// --- Siemens Structured Format ---
DATA_BLOCK "model__HS8_IW50_"
{ S7_Optimized_Access := 'TRUE' }
VERSION :
NON_RETAIN
   VAR
      W_i : ARRAY[0..7, 0..39] OF REAL;
      W_f : ARRAY[0..7, 0..39] OF REAL;
      W_g : ARRAY[0..7, 0..39] OF REAL;
      W_o : ARRAY[0..7, 0..39] OF REAL;
      R_i : ARRAY[0..7, 0..7] OF REAL;
      R_f : ARRAY[0..7, 0..7] OF REAL;
      R_g : ARRAY[0..7, 0..7] OF REAL;
      R_o : ARRAY[0..7, 0..7] OF REAL;
      B_i : ARRAY[0..7] OF REAL;
      B_f : ARRAY[0..7] OF REAL;
      B_g : ARRAY[0..7] OF REAL;
      B_o : ARRAY[0..7] OF REAL;
      FC_W : ARRAY[0..39, 0..7] OF REAL;
      FC_B : ARRAY[0..39] OF REAL;
   END_VAR
BEGIN

      W_i[0,0] := 0.02461717;
      W_i[0,1] := 0.08401545;
      W_i[0,2] := -0.12303820;
      W_i[0,3] := -0.02682650;
      W_i[0,4] := 0.14538512;
      W_i[0,5] := 0.05910228;
      W_i[0,6] := -0.06121323;
      W_i[0,7] := 0.19529903;
      W_i[0,8] := 0.21199454;
      W_i[0,9] := -0.29979098;
      W_i[0,10] := -0.09429822;
      W_i[0,11] := -0.28532824;
      W_i[0,12] := 0.06377743;
      W_i[0,13] := -0.06364888;
      W_i[0,14] := 0.00534459;
      W_i[0,15] := 0.03598412;
      W_i[0,16] := 0.04236616;
      W_i[0,17] := 0.00850482;
      W_i[0,18] := 0.00358703;
      W_i[0,19] := 0.18395557;
      W_i[0,20] := 0.05710260;
      W_i[0,21] := 0.31176916;
      W_i[0,22] := 0.17010060;
      W_i[0,23] := -0.01221133;
      W_i[0,24] := -0.19286193;
      W_i[0,25] := -0.07674938;
      W_i[0,26] := -0.40142074;
      W_i[0,27] := -0.50435519;
      W_i[0,28] := 0.04934237;
      W_i[0,29] := -0.24499206;
      W_i[0,30] := 0.63579166;
      W_i[0,31] := -0.13499857;
      W_i[0,32] := 0.02890123;
      W_i[0,33] := -0.00438442;
      W_i[0,34] := -0.02304220;
      W_i[0,35] := -0.28221473;
      W_i[0,36] := -0.00601982;
      W_i[0,37] := -0.39292136;
      W_i[0,38] := -0.02013459;
      W_i[0,39] := -0.00859181;
      W_i[1,0] := -0.17783616;
      W_i[1,1] := 0.10906062;
      W_i[1,2] := 0.27302170;
      W_i[1,3] := 0.03857158;
      W_i[1,4] := 0.15132146;
      W_i[1,5] := -0.07943013;
      W_i[1,6] := -0.12445311;
      W_i[1,7] := 0.10142804;
      W_i[1,8] := 0.17782561;
      W_i[1,9] := -0.34472182;
      W_i[1,10] := -0.15930130;
      W_i[1,11] := 0.11785957;
      W_i[1,12] := 0.12351760;
      W_i[1,13] := 0.01896391;
      W_i[1,14] := -0.06655354;
      W_i[1,15] := 0.10417320;
      W_i[1,16] := 0.02300226;
      W_i[1,17] := -0.06141837;
      W_i[1,18] := 0.28663757;
      W_i[1,19] := -0.05906216;
      W_i[1,20] := -0.01470305;
      W_i[1,21] := 0.12249159;
      W_i[1,22] := 0.08935670;
      W_i[1,23] := -0.19675028;
      W_i[1,24] := 0.48150146;
      W_i[1,25] := 0.29962191;
      W_i[1,26] := 0.04253698;
      W_i[1,27] := -0.01234774;
      W_i[1,28] := -0.20131898;
      W_i[1,29] := -0.28958127;
      W_i[1,30] := 0.30615368;
      W_i[1,31] := -0.00297963;
      W_i[1,32] := 0.24898766;
      W_i[1,33] := -0.17079352;
      W_i[1,34] := -0.01789305;
      W_i[1,35] := -0.07885017;
      W_i[1,36] := 0.02689386;
      W_i[1,37] := 0.36441922;
      W_i[1,38] := -0.06345996;
      W_i[1,39] := 0.09888364;
      W_i[2,0] := 0.10794700;
      W_i[2,1] := 0.01449859;
      W_i[2,2] := 0.11232290;
      W_i[2,3] := 0.04600843;
      W_i[2,4] := 0.15555517;
      W_i[2,5] := -0.08419870;
      W_i[2,6] := 0.10784180;
      W_i[2,7] := -0.13110802;
      W_i[2,8] := 0.01003856;
      W_i[2,9] := 0.13528554;
      W_i[2,10] := -0.08593279;
      W_i[2,11] := 0.15705661;
      W_i[2,12] := 0.00744481;
      W_i[2,13] := 0.14232995;
      W_i[2,14] := -0.07310586;
      W_i[2,15] := 0.11869515;
      W_i[2,16] := 0.16272350;
      W_i[2,17] := 0.01258006;
      W_i[2,18] := 0.17897964;
      W_i[2,19] := -0.08531563;
      W_i[2,20] := -0.06869420;
      W_i[2,21] := -0.05605607;
      W_i[2,22] := -0.24934621;
      W_i[2,23] := 0.02436493;
      W_i[2,24] := 0.04889333;
      W_i[2,25] := -0.20094825;
      W_i[2,26] := -0.40725628;
      W_i[2,27] := -0.16053441;
      W_i[2,28] := -0.17641398;
      W_i[2,29] := -0.18513416;
      W_i[2,30] := 0.09812243;
      W_i[2,31] := -0.24586804;
      W_i[2,32] := 0.18386346;
      W_i[2,33] := -0.37200448;
      W_i[2,34] := -0.30738470;
      W_i[2,35] := 0.07613509;
      W_i[2,36] := -0.04531293;
      W_i[2,37] := -0.08632755;
      W_i[2,38] := -0.13347539;
      W_i[2,39] := -0.03515237;
      W_i[3,0] := -0.04817922;
      W_i[3,1] := -0.16765678;
      W_i[3,2] := -0.00308369;
      W_i[3,3] := -0.41362956;
      W_i[3,4] := -0.07394656;
      W_i[3,5] := 0.09627691;
      W_i[3,6] := 0.11941688;
      W_i[3,7] := -0.17643057;
      W_i[3,8] := 0.06146013;
      W_i[3,9] := 0.13595612;
      W_i[3,10] := 0.21689560;
      W_i[3,11] := 0.08097983;
      W_i[3,12] := -0.05968216;
      W_i[3,13] := 0.06028462;
      W_i[3,14] := -0.33660558;
      W_i[3,15] := -0.14613369;
      W_i[3,16] := 0.15110187;
      W_i[3,17] := 0.02597690;
      W_i[3,18] := 0.00098816;
      W_i[3,19] := 0.26554033;
      W_i[3,20] := 0.06123941;
      W_i[3,21] := -0.20589893;
      W_i[3,22] := -0.01046670;
      W_i[3,23] := -0.35783783;
      W_i[3,24] := -0.18957515;
      W_i[3,25] := -0.03140980;
      W_i[3,26] := 0.00826861;
      W_i[3,27] := 0.05130741;
      W_i[3,28] := 0.13812958;
      W_i[3,29] := -0.19599199;
      W_i[3,30] := -0.16747603;
      W_i[3,31] := -0.13670678;
      W_i[3,32] := -0.15334715;
      W_i[3,33] := -0.32899481;
      W_i[3,34] := 0.07909799;
      W_i[3,35] := -0.27765223;
      W_i[3,36] := -0.03015585;
      W_i[3,37] := 0.07159591;
      W_i[3,38] := -0.33855185;
      W_i[3,39] := -0.69761050;
      W_i[4,0] := 0.10504181;
      W_i[4,1] := 0.00682971;
      W_i[4,2] := -0.05512364;
      W_i[4,3] := -0.42238507;
      W_i[4,4] := 0.21000206;
      W_i[4,5] := 0.08828816;
      W_i[4,6] := -0.25787413;
      W_i[4,7] := 0.18548162;
      W_i[4,8] := 0.07325415;
      W_i[4,9] := -0.16746196;
      W_i[4,10] := -0.23054802;
      W_i[4,11] := -0.17278661;
      W_i[4,12] := 0.19685929;
      W_i[4,13] := -0.06621253;
      W_i[4,14] := -0.04979985;
      W_i[4,15] := -0.02534566;
      W_i[4,16] := -0.05196558;
      W_i[4,17] := -0.02844546;
      W_i[4,18] := 0.21438381;
      W_i[4,19] := -0.22215076;
      W_i[4,20] := 0.01178194;
      W_i[4,21] := -0.06624336;
      W_i[4,22] := -0.05115673;
      W_i[4,23] := -0.23732296;
      W_i[4,24] := -0.09036870;
      W_i[4,25] := -0.09140033;
      W_i[4,26] := 0.12307051;
      W_i[4,27] := -0.02017660;
      W_i[4,28] := -0.07642211;
      W_i[4,29] := -0.01614011;
      W_i[4,30] := -0.17466348;
      W_i[4,31] := -0.15838575;
      W_i[4,32] := 0.18079966;
      W_i[4,33] := 0.33373138;
      W_i[4,34] := 0.09327173;
      W_i[4,35] := -0.13638979;
      W_i[4,36] := -0.08043678;
      W_i[4,37] := -0.09420969;
      W_i[4,38] := -0.03976285;
      W_i[4,39] := 0.22526605;
      W_i[5,0] := 0.46471885;
      W_i[5,1] := 0.24254853;
      W_i[5,2] := -0.00896330;
      W_i[5,3] := -0.40931293;
      W_i[5,4] := 0.07764716;
      W_i[5,5] := -0.12571707;
      W_i[5,6] := -0.07207277;
      W_i[5,7] := -0.58136684;
      W_i[5,8] := -0.70827621;
      W_i[5,9] := 0.13912673;
      W_i[5,10] := 0.00305168;
      W_i[5,11] := 0.10330518;
      W_i[5,12] := -0.39406857;
      W_i[5,13] := -0.13641670;
      W_i[5,14] := -0.13437758;
      W_i[5,15] := 0.32282859;
      W_i[5,16] := 0.14888868;
      W_i[5,17] := 0.07580157;
      W_i[5,18] := 0.78602076;
      W_i[5,19] := -0.46361649;
      W_i[5,20] := -0.12363275;
      W_i[5,21] := 0.16991106;
      W_i[5,22] := -0.08441558;
      W_i[5,23] := 0.01862625;
      W_i[5,24] := 0.45371729;
      W_i[5,25] := 1.03232503;
      W_i[5,26] := 0.00888214;
      W_i[5,27] := -0.04149527;
      W_i[5,28] := -0.06423787;
      W_i[5,29] := -0.13104723;
      W_i[5,30] := -0.16760458;
      W_i[5,31] := -0.06425823;
      W_i[5,32] := 0.11957818;
      W_i[5,33] := 0.10409375;
      W_i[5,34] := 0.68515724;
      W_i[5,35] := 0.21046008;
      W_i[5,36] := 0.09369295;
      W_i[5,37] := -0.08919100;
      W_i[5,38] := -0.09835245;
      W_i[5,39] := 0.00684949;
      W_i[6,0] := 0.04514975;
      W_i[6,1] := -0.18210933;
      W_i[6,2] := -0.00654514;
      W_i[6,3] := -0.41125798;
      W_i[6,4] := 0.04396775;
      W_i[6,5] := -0.00702968;
      W_i[6,6] := -0.05002901;
      W_i[6,7] := -0.03861308;
      W_i[6,8] := 0.06189432;
      W_i[6,9] := -0.02187389;
      W_i[6,10] := 0.03767673;
      W_i[6,11] := -0.55604023;
      W_i[6,12] := -0.48857787;
      W_i[6,13] := 0.13115734;
      W_i[6,14] := -0.05613643;
      W_i[6,15] := -0.11288932;
      W_i[6,16] := 0.17460676;
      W_i[6,17] := -0.26465502;
      W_i[6,18] := 0.16549894;
      W_i[6,19] := 0.29697806;
      W_i[6,20] := 0.23571719;
      W_i[6,21] := -0.09589785;
      W_i[6,22] := 0.59926170;
      W_i[6,23] := -0.08488554;
      W_i[6,24] := 0.70308256;
      W_i[6,25] := 0.90409851;
      W_i[6,26] := -0.01121288;
      W_i[6,27] := -0.09806376;
      W_i[6,28] := -0.02374482;
      W_i[6,29] := -0.20431902;
      W_i[6,30] := 0.48442781;
      W_i[6,31] := -0.11867638;
      W_i[6,32] := 0.28192973;
      W_i[6,33] := 0.13702093;
      W_i[6,34] := 0.91159022;
      W_i[6,35] := -0.05850424;
      W_i[6,36] := -0.02443852;
      W_i[6,37] := 0.08158594;
      W_i[6,38] := -0.16384257;
      W_i[6,39] := 0.04486246;
      W_i[7,0] := -0.16619515;
      W_i[7,1] := -0.08064937;
      W_i[7,2] := 0.17380525;
      W_i[7,3] := -0.35741210;
      W_i[7,4] := 0.25576842;
      W_i[7,5] := -0.11047508;
      W_i[7,6] := -0.00358257;
      W_i[7,7] := 0.22714809;
      W_i[7,8] := 0.14583488;
      W_i[7,9] := -0.14972806;
      W_i[7,10] := -0.14519584;
      W_i[7,11] := -0.41559315;
      W_i[7,12] := -0.01696615;
      W_i[7,13] := -0.28414848;
      W_i[7,14] := 0.06566004;
      W_i[7,15] := 0.09450804;
      W_i[7,16] := -0.03949518;
      W_i[7,17] := 0.04709280;
      W_i[7,18] := 0.19348225;
      W_i[7,19] := 0.10500827;
      W_i[7,20] := -0.09005301;
      W_i[7,21] := -0.34911180;
      W_i[7,22] := -0.00604367;
      W_i[7,23] := -0.15790336;
      W_i[7,24] := 0.51519841;
      W_i[7,25] := 1.09936786;
      W_i[7,26] := -0.23214035;
      W_i[7,27] := -0.30644259;
      W_i[7,28] := 0.08868466;
      W_i[7,29] := 0.18681195;
      W_i[7,30] := 0.44118169;
      W_i[7,31] := 0.16998404;
      W_i[7,32] := -0.39800110;
      W_i[7,33] := 0.02014814;
      W_i[7,34] := 0.50454497;
      W_i[7,35] := -0.04675045;
      W_i[7,36] := -0.05744690;
      W_i[7,37] := 0.17443271;
      W_i[7,38] := -0.05675455;
      W_i[7,39] := 0.18483149;
      W_f[0,0] := -0.08831103;
      W_f[0,1] := 0.00681163;
      W_f[0,2] := -0.02927266;
      W_f[0,3] := 0.05481192;
      W_f[0,4] := -0.06411999;
      W_f[0,5] := 0.00323826;
      W_f[0,6] := 0.04202358;
      W_f[0,7] := -0.14036146;
      W_f[0,8] := -0.12626842;
      W_f[0,9] := 0.10009770;
      W_f[0,10] := 0.02791548;
      W_f[0,11] := -0.04096280;
      W_f[0,12] := -0.00354303;
      W_f[0,13] := 0.01158499;
      W_f[0,14] := -0.04464640;
      W_f[0,15] := -0.08357976;
      W_f[0,16] := 0.04911109;
      W_f[0,17] := 0.09140756;
      W_f[0,18] := -0.03252059;
      W_f[0,19] := 0.01830712;
      W_f[0,20] := 0.01689613;
      W_f[0,21] := 0.22018659;
      W_f[0,22] := 0.08402620;
      W_f[0,23] := -0.07398796;
      W_f[0,24] := 0.08441300;
      W_f[0,25] := 0.18096766;
      W_f[0,26] := 0.05508868;
      W_f[0,27] := -0.13029598;
      W_f[0,28] := -0.02453627;
      W_f[0,29] := 0.12306897;
      W_f[0,30] := 0.37074596;
      W_f[0,31] := 0.04067184;
      W_f[0,32] := 0.33210105;
      W_f[0,33] := 0.17263570;
      W_f[0,34] := 0.02185974;
      W_f[0,35] := 0.21439323;
      W_f[0,36] := 0.00803035;
      W_f[0,37] := 0.09185252;
      W_f[0,38] := -0.03025025;
      W_f[0,39] := 0.16901997;
      W_f[1,0] := -0.08017771;
      W_f[1,1] := 0.05072340;
      W_f[1,2] := -0.15171054;
      W_f[1,3] := -0.04507771;
      W_f[1,4] := -0.01952654;
      W_f[1,5] := 0.01524715;
      W_f[1,6] := -0.03147047;
      W_f[1,7] := -0.02802088;
      W_f[1,8] := -0.15045448;
      W_f[1,9] := 0.13191310;
      W_f[1,10] := 0.00395375;
      W_f[1,11] := -0.03943809;
      W_f[1,12] := -0.13766901;
      W_f[1,13] := -0.04960233;
      W_f[1,14] := -0.11882943;
      W_f[1,15] := -0.18921053;
      W_f[1,16] := 0.07628337;
      W_f[1,17] := -0.01504870;
      W_f[1,18] := 0.23253591;
      W_f[1,19] := 0.00738192;
      W_f[1,20] := 0.02966039;
      W_f[1,21] := -0.07575663;
      W_f[1,22] := 0.28070211;
      W_f[1,23] := 0.04504234;
      W_f[1,24] := 0.44733906;
      W_f[1,25] := 0.76406956;
      W_f[1,26] := -0.18153259;
      W_f[1,27] := -0.01630468;
      W_f[1,28] := 0.04244527;
      W_f[1,29] := -0.03562038;
      W_f[1,30] := 0.06799272;
      W_f[1,31] := -0.07704592;
      W_f[1,32] := 0.08059093;
      W_f[1,33] := 0.21711972;
      W_f[1,34] := 0.58922273;
      W_f[1,35] := -0.24995837;
      W_f[1,36] := -0.01296289;
      W_f[1,37] := -0.02005322;
      W_f[1,38] := 0.11887441;
      W_f[1,39] := 0.13964133;
      W_f[2,0] := 0.02022752;
      W_f[2,1] := -0.03258032;
      W_f[2,2] := 0.02105030;
      W_f[2,3] := -0.01033732;
      W_f[2,4] := -0.02927784;
      W_f[2,5] := 0.05956579;
      W_f[2,6] := -0.06668916;
      W_f[2,7] := -0.06423724;
      W_f[2,8] := -0.06636658;
      W_f[2,9] := 0.16499053;
      W_f[2,10] := -0.01066389;
      W_f[2,11] := -0.08655350;
      W_f[2,12] := 0.03831896;
      W_f[2,13] := 0.02458346;
      W_f[2,14] := 0.12203392;
      W_f[2,15] := -0.07686506;
      W_f[2,16] := -0.09261417;
      W_f[2,17] := -0.01410419;
      W_f[2,18] := 0.05016823;
      W_f[2,19] := -0.13551356;
      W_f[2,20] := 0.00147612;
      W_f[2,21] := -0.01080879;
      W_f[2,22] := -0.23093474;
      W_f[2,23] := 0.18362746;
      W_f[2,24] := 0.34206459;
      W_f[2,25] := 0.11531623;
      W_f[2,26] := -0.10813569;
      W_f[2,27] := -0.03727976;
      W_f[2,28] := 0.08597951;
      W_f[2,29] := 0.16925062;
      W_f[2,30] := 0.14001821;
      W_f[2,31] := 0.08336479;
      W_f[2,32] := -0.13725568;
      W_f[2,33] := 0.14078599;
      W_f[2,34] := -0.22189134;
      W_f[2,35] := 0.07339284;
      W_f[2,36] := 0.01494332;
      W_f[2,37] := -0.16808337;
      W_f[2,38] := 0.02411579;
      W_f[2,39] := 0.21152344;
      W_f[3,0] := -0.03794771;
      W_f[3,1] := 0.05475021;
      W_f[3,2] := -0.02614000;
      W_f[3,3] := 0.08930103;
      W_f[3,4] := 0.04492093;
      W_f[3,5] := 0.03020424;
      W_f[3,6] := -0.07041149;
      W_f[3,7] := 0.23536491;
      W_f[3,8] := -0.04178810;
      W_f[3,9] := -0.19159153;
      W_f[3,10] := -0.06868339;
      W_f[3,11] := -0.16539882;
      W_f[3,12] := 0.12754864;
      W_f[3,13] := -0.13497283;
      W_f[3,14] := 0.13930795;
      W_f[3,15] := 0.00134255;
      W_f[3,16] := -0.03635018;
      W_f[3,17] := 0.02573154;
      W_f[3,18] := -0.41695386;
      W_f[3,19] := -0.18809830;
      W_f[3,20] := 0.04352702;
      W_f[3,21] := 0.16437882;
      W_f[3,22] := 0.06266205;
      W_f[3,23] := 0.08159398;
      W_f[3,24] := 0.04201810;
      W_f[3,25] := -0.19031751;
      W_f[3,26] := -0.17173289;
      W_f[3,27] := -0.23532763;
      W_f[3,28] := 0.17517763;
      W_f[3,29] := 0.39156693;
      W_f[3,30] := 0.25430456;
      W_f[3,31] := 0.07574216;
      W_f[3,32] := 0.27996075;
      W_f[3,33] := 0.00114326;
      W_f[3,34] := -0.28795609;
      W_f[3,35] := 0.19662365;
      W_f[3,36] := 0.02395431;
      W_f[3,37] := -0.22338727;
      W_f[3,38] := 0.15306281;
      W_f[3,39] := 0.18428560;
      W_f[4,0] := 0.01311270;
      W_f[4,1] := -0.01359527;
      W_f[4,2] := -0.03426387;
      W_f[4,3] := -0.05035185;
      W_f[4,4] := 0.09912422;
      W_f[4,5] := -0.04895325;
      W_f[4,6] := -0.03395505;
      W_f[4,7] := -0.02843624;
      W_f[4,8] := -0.08145776;
      W_f[4,9] := 0.08917268;
      W_f[4,10] := -0.00391436;
      W_f[4,11] := -0.07863925;
      W_f[4,12] := 0.03092329;
      W_f[4,13] := 0.01714266;
      W_f[4,14] := -0.03228388;
      W_f[4,15] := -0.05111328;
      W_f[4,16] := 0.02532922;
      W_f[4,17] := -0.04550080;
      W_f[4,18] := -0.03456742;
      W_f[4,19] := -0.02089478;
      W_f[4,20] := 0.09678645;
      W_f[4,21] := -0.08640780;
      W_f[4,22] := 0.02293069;
      W_f[4,23] := 0.05295998;
      W_f[4,24] := 0.11747785;
      W_f[4,25] := 0.00186043;
      W_f[4,26] := -0.20221773;
      W_f[4,27] := -0.01488341;
      W_f[4,28] := 0.04745471;
      W_f[4,29] := -0.16965286;
      W_f[4,30] := 0.02288965;
      W_f[4,31] := -0.03804171;
      W_f[4,32] := 0.13254493;
      W_f[4,33] := -0.13787529;
      W_f[4,34] := -0.43391764;
      W_f[4,35] := -0.24835001;
      W_f[4,36] := 0.07141465;
      W_f[4,37] := -0.29939890;
      W_f[4,38] := -0.01851079;
      W_f[4,39] := 0.08986987;
      W_f[5,0] := -0.14319988;
      W_f[5,1] := -0.10292582;
      W_f[5,2] := -0.17382213;
      W_f[5,3] := -0.01608473;
      W_f[5,4] := -0.00378885;
      W_f[5,5] := 0.00846169;
      W_f[5,6] := 0.06387471;
      W_f[5,7] := 0.20796628;
      W_f[5,8] := -0.42914653;
      W_f[5,9] := 0.01919760;
      W_f[5,10] := 0.04385304;
      W_f[5,11] := 0.01982332;
      W_f[5,12] := 0.11683133;
      W_f[5,13] := 0.07871818;
      W_f[5,14] := -0.12016966;
      W_f[5,15] := -0.06522254;
      W_f[5,16] := -0.10883621;
      W_f[5,17] := -0.02835156;
      W_f[5,18] := -0.26717833;
      W_f[5,19] := 0.08458684;
      W_f[5,20] := -0.00364884;
      W_f[5,21] := -0.04485849;
      W_f[5,22] := -0.19082835;
      W_f[5,23] := 0.06622007;
      W_f[5,24] := 0.45456037;
      W_f[5,25] := 0.15541779;
      W_f[5,26] := 0.00758505;
      W_f[5,27] := 0.07440008;
      W_f[5,28] := 0.05810034;
      W_f[5,29] := 0.14797372;
      W_f[5,30] := -0.11548296;
      W_f[5,31] := 0.02787589;
      W_f[5,32] := -0.27752876;
      W_f[5,33] := -0.08107541;
      W_f[5,34] := -0.09626248;
      W_f[5,35] := -0.23543228;
      W_f[5,36] := -0.00549724;
      W_f[5,37] := 0.06302677;
      W_f[5,38] := 0.14402032;
      W_f[5,39] := 0.31771937;
      W_f[6,0] := 0.05912529;
      W_f[6,1] := 0.00633830;
      W_f[6,2] := -0.00901835;
      W_f[6,3] := -0.10450855;
      W_f[6,4] := 0.03491682;
      W_f[6,5] := 0.04512391;
      W_f[6,6] := 0.04958262;
      W_f[6,7] := 0.01803463;
      W_f[6,8] := -0.04358606;
      W_f[6,9] := -0.09593592;
      W_f[6,10] := 0.00282181;
      W_f[6,11] := -0.14376016;
      W_f[6,12] := 0.10038611;
      W_f[6,13] := -0.04489579;
      W_f[6,14] := 0.06795548;
      W_f[6,15] := -0.00965744;
      W_f[6,16] := 0.03404293;
      W_f[6,17] := 0.02229516;
      W_f[6,18] := -0.14460719;
      W_f[6,19] := -0.22980542;
      W_f[6,20] := 0.11291888;
      W_f[6,21] := 0.08677951;
      W_f[6,22] := 0.57823741;
      W_f[6,23] := 0.01069405;
      W_f[6,24] := 0.79735392;
      W_f[6,25] := 0.83291894;
      W_f[6,26] := 0.03028462;
      W_f[6,27] := -0.03470038;
      W_f[6,28] := 0.03831891;
      W_f[6,29] := -0.38390651;
      W_f[6,30] := 0.59899300;
      W_f[6,31] := 0.08223967;
      W_f[6,32] := 0.27525041;
      W_f[6,33] := 0.50554472;
      W_f[6,34] := 0.56139988;
      W_f[6,35] := 0.04573379;
      W_f[6,36] := -0.01382815;
      W_f[6,37] := -0.07028573;
      W_f[6,38] := 0.02817321;
      W_f[6,39] := 0.01610095;
      W_f[7,0] := -0.00575910;
      W_f[7,1] := 0.01253089;
      W_f[7,2] := -0.03966596;
      W_f[7,3] := -0.04416019;
      W_f[7,4] := -0.04916450;
      W_f[7,5] := 0.00926291;
      W_f[7,6] := -0.00996001;
      W_f[7,7] := -0.06242750;
      W_f[7,8] := -0.03272317;
      W_f[7,9] := 0.14268650;
      W_f[7,10] := 0.00977653;
      W_f[7,11] := -0.17324640;
      W_f[7,12] := -0.05803645;
      W_f[7,13] := -0.05088602;
      W_f[7,14] := 0.00851257;
      W_f[7,15] := -0.08858407;
      W_f[7,16] := 0.11187664;
      W_f[7,17] := -0.00764770;
      W_f[7,18] := 0.13751905;
      W_f[7,19] := 0.15364748;
      W_f[7,20] := 0.01291497;
      W_f[7,21] := 0.08050860;
      W_f[7,22] := 0.02860431;
      W_f[7,23] := 0.02334928;
      W_f[7,24] := 0.27481839;
      W_f[7,25] := 0.06242412;
      W_f[7,26] := -0.03117798;
      W_f[7,27] := -0.06928296;
      W_f[7,28] := -0.02172423;
      W_f[7,29] := 0.26392910;
      W_f[7,30] := 0.09593272;
      W_f[7,31] := -0.05563883;
      W_f[7,32] := 0.16712280;
      W_f[7,33] := 0.18572508;
      W_f[7,34] := 0.03861195;
      W_f[7,35] := -0.06280123;
      W_f[7,36] := -0.00801319;
      W_f[7,37] := -0.12490637;
      W_f[7,38] := -0.14012046;
      W_f[7,39] := 0.13752492;
      W_g[0,0] := -0.05256320;
      W_g[0,1] := 0.03376590;
      W_g[0,2] := -0.05004627;
      W_g[0,3] := 0.01062740;
      W_g[0,4] := -0.17505662;
      W_g[0,5] := 0.04523542;
      W_g[0,6] := 0.10033184;
      W_g[0,7] := 0.01237159;
      W_g[0,8] := 0.00997229;
      W_g[0,9] := 0.01509623;
      W_g[0,10] := -0.03384563;
      W_g[0,11] := 0.01027409;
      W_g[0,12] := 0.01079937;
      W_g[0,13] := -0.00604036;
      W_g[0,14] := -0.05007736;
      W_g[0,15] := -0.01323667;
      W_g[0,16] := 0.01487322;
      W_g[0,17] := 0.10829928;
      W_g[0,18] := -0.01920407;
      W_g[0,19] := 0.01481452;
      W_g[0,20] := -0.10726670;
      W_g[0,21] := 0.10591213;
      W_g[0,22] := -0.06350547;
      W_g[0,23] := -0.00731946;
      W_g[0,24] := 0.19152513;
      W_g[0,25] := 0.07594201;
      W_g[0,26] := -0.05230021;
      W_g[0,27] := 0.15840378;
      W_g[0,28] := -0.11106505;
      W_g[0,29] := -0.00231445;
      W_g[0,30] := 0.03844558;
      W_g[0,31] := 0.00872381;
      W_g[0,32] := -0.03187981;
      W_g[0,33] := 0.00040774;
      W_g[0,34] := -0.19478397;
      W_g[0,35] := 0.15274970;
      W_g[0,36] := 0.02823638;
      W_g[0,37] := -0.10759887;
      W_g[0,38] := -0.04167965;
      W_g[0,39] := -0.03888805;
      W_g[1,0] := -0.08446153;
      W_g[1,1] := 0.05808212;
      W_g[1,2] := -0.08208533;
      W_g[1,3] := 0.03618253;
      W_g[1,4] := -0.05700465;
      W_g[1,5] := 0.02161270;
      W_g[1,6] := -0.00616194;
      W_g[1,7] := 0.02231257;
      W_g[1,8] := 0.02348651;
      W_g[1,9] := 0.00478895;
      W_g[1,10] := 0.03830986;
      W_g[1,11] := 0.13621216;
      W_g[1,12] := 0.11095273;
      W_g[1,13] := 0.01325371;
      W_g[1,14] := -0.01293219;
      W_g[1,15] := 0.12523465;
      W_g[1,16] := -0.06386022;
      W_g[1,17] := -0.06564955;
      W_g[1,18] := -0.07677279;
      W_g[1,19] := 0.13738941;
      W_g[1,20] := 0.00232198;
      W_g[1,21] := -0.04238968;
      W_g[1,22] := -0.06318325;
      W_g[1,23] := 0.03427328;
      W_g[1,24] := 0.18657008;
      W_g[1,25] := -0.18876043;
      W_g[1,26] := 0.04970511;
      W_g[1,27] := -0.04672737;
      W_g[1,28] := -0.03255373;
      W_g[1,29] := 0.00354951;
      W_g[1,30] := 0.06089024;
      W_g[1,31] := 0.00000845;
      W_g[1,32] := 0.00405714;
      W_g[1,33] := -0.01229481;
      W_g[1,34] := 0.42297170;
      W_g[1,35] := 0.32250756;
      W_g[1,36] := -0.04902744;
      W_g[1,37] := -0.30256015;
      W_g[1,38] := -0.03282990;
      W_g[1,39] := -0.03006732;
      W_g[2,0] := 0.08679828;
      W_g[2,1] := -0.01636712;
      W_g[2,2] := 0.08163529;
      W_g[2,3] := 0.04131987;
      W_g[2,4] := -0.12495904;
      W_g[2,5] := 0.04998558;
      W_g[2,6] := 0.05360224;
      W_g[2,7] := 0.00646355;
      W_g[2,8] := 0.01505343;
      W_g[2,9] := 0.03555880;
      W_g[2,10] := 0.01924760;
      W_g[2,11] := -0.02805754;
      W_g[2,12] := -0.02042336;
      W_g[2,13] := 0.11497736;
      W_g[2,14] := 0.02289071;
      W_g[2,15] := -0.00648216;
      W_g[2,16] := 0.00574631;
      W_g[2,17] := -0.03994992;
      W_g[2,18] := -0.10415535;
      W_g[2,19] := 0.01829612;
      W_g[2,20] := -0.05056486;
      W_g[2,21] := 0.02768292;
      W_g[2,22] := 0.01188622;
      W_g[2,23] := 0.12093837;
      W_g[2,24] := -0.00732198;
      W_g[2,25] := 0.06027466;
      W_g[2,26] := 0.06612495;
      W_g[2,27] := 0.00363937;
      W_g[2,28] := -0.05205845;
      W_g[2,29] := -0.08297625;
      W_g[2,30] := -0.00665878;
      W_g[2,31] := 0.01979631;
      W_g[2,32] := -0.00752764;
      W_g[2,33] := -0.00295640;
      W_g[2,34] := 0.54437882;
      W_g[2,35] := -0.15383327;
      W_g[2,36] := -0.03264818;
      W_g[2,37] := 0.17412139;
      W_g[2,38] := 0.05972110;
      W_g[2,39] := 0.04769525;
      W_g[3,0] := 0.05698530;
      W_g[3,1] := -0.00717941;
      W_g[3,2] := 0.06096774;
      W_g[3,3] := -0.04463135;
      W_g[3,4] := -0.13414808;
      W_g[3,5] := -0.04385218;
      W_g[3,6] := -0.09330478;
      W_g[3,7] := -0.06749506;
      W_g[3,8] := -0.05428461;
      W_g[3,9] := -0.02963200;
      W_g[3,10] := 0.00547227;
      W_g[3,11] := -0.05570020;
      W_g[3,12] := -0.04208678;
      W_g[3,13] := 0.03579268;
      W_g[3,14] := 0.02666621;
      W_g[3,15] := -0.01365136;
      W_g[3,16] := -0.03459660;
      W_g[3,17] := -0.11479730;
      W_g[3,18] := -0.05903023;
      W_g[3,19] := -0.05609168;
      W_g[3,20] := 0.06238525;
      W_g[3,21] := 0.04947945;
      W_g[3,22] := 0.04299555;
      W_g[3,23] := 0.03366689;
      W_g[3,24] := -0.47512600;
      W_g[3,25] := -0.63947034;
      W_g[3,26] := -0.05774437;
      W_g[3,27] := 0.06282470;
      W_g[3,28] := -0.15790993;
      W_g[3,29] := 0.20147590;
      W_g[3,30] := -0.11538504;
      W_g[3,31] := -0.01063631;
      W_g[3,32] := 0.00111993;
      W_g[3,33] := -0.01895600;
      W_g[3,34] := -0.15655167;
      W_g[3,35] := -0.16384147;
      W_g[3,36] := 0.04147036;
      W_g[3,37] := 0.13167211;
      W_g[3,38] := 0.02300073;
      W_g[3,39] := 0.42263514;
      W_g[4,0] := -0.01835994;
      W_g[4,1] := -0.01981971;
      W_g[4,2] := -0.01484892;
      W_g[4,3] := 0.04219592;
      W_g[4,4] := -0.03390066;
      W_g[4,5] := 0.05298800;
      W_g[4,6] := 0.08669198;
      W_g[4,7] := 0.07381222;
      W_g[4,8] := 0.05830150;
      W_g[4,9] := 0.04904483;
      W_g[4,10] := 0.01153296;
      W_g[4,11] := 0.00024178;
      W_g[4,12] := 0.01480092;
      W_g[4,13] := -0.01464547;
      W_g[4,14] := 0.03931813;
      W_g[4,15] := -0.00775862;
      W_g[4,16] := 0.07005515;
      W_g[4,17] := 0.07610738;
      W_g[4,18] := -0.06145393;
      W_g[4,19] := 0.01960655;
      W_g[4,20] := -0.08848560;
      W_g[4,21] := -0.01328403;
      W_g[4,22] := -0.12893535;
      W_g[4,23] := 0.01238164;
      W_g[4,24] := -0.43381751;
      W_g[4,25] := -0.31650203;
      W_g[4,26] := -0.00358412;
      W_g[4,27] := -0.00217345;
      W_g[4,28] := 0.03488368;
      W_g[4,29] := -0.06516429;
      W_g[4,30] := 0.03693077;
      W_g[4,31] := -0.03261345;
      W_g[4,32] := -0.07810706;
      W_g[4,33] := -0.06320744;
      W_g[4,34] := -0.11921121;
      W_g[4,35] := 0.02571805;
      W_g[4,36] := -0.06975383;
      W_g[4,37] := -0.13379739;
      W_g[4,38] := 0.04367201;
      W_g[4,39] := 0.03239072;
      W_g[5,0] := 0.20069297;
      W_g[5,1] := -0.16023712;
      W_g[5,2] := 0.17268215;
      W_g[5,3] := 0.09593190;
      W_g[5,4] := -0.00601159;
      W_g[5,5] := -0.05667128;
      W_g[5,6] := -0.02598925;
      W_g[5,7] := 0.06759191;
      W_g[5,8] := 0.04750817;
      W_g[5,9] := 0.21007423;
      W_g[5,10] := 0.09670225;
      W_g[5,11] := -0.02642447;
      W_g[5,12] := 0.01532454;
      W_g[5,13] := 0.01303505;
      W_g[5,14] := -0.08846440;
      W_g[5,15] := 0.01258479;
      W_g[5,16] := -0.04598146;
      W_g[5,17] := -0.03127987;
      W_g[5,18] := 0.47458670;
      W_g[5,19] := -0.00303655;
      W_g[5,20] := 0.02677378;
      W_g[5,21] := 0.02378645;
      W_g[5,22] := 0.03294978;
      W_g[5,23] := 0.05323023;
      W_g[5,24] := -0.08479793;
      W_g[5,25] := 0.37677112;
      W_g[5,26] := -0.02968354;
      W_g[5,27] := 0.02218193;
      W_g[5,28] := -0.00680012;
      W_g[5,29] := -0.02114836;
      W_g[5,30] := -0.03917154;
      W_g[5,31] := -0.01134670;
      W_g[5,32] := -0.00775183;
      W_g[5,33] := -0.01060248;
      W_g[5,34] := 0.13405052;
      W_g[5,35] := -0.07177506;
      W_g[5,36] := 0.02046018;
      W_g[5,37] := 0.04711805;
      W_g[5,38] := -0.09608429;
      W_g[5,39] := -0.06293187;
      W_g[6,0] := 0.05725823;
      W_g[6,1] := -0.01282716;
      W_g[6,2] := 0.05448377;
      W_g[6,3] := -0.04432564;
      W_g[6,4] := 0.02756098;
      W_g[6,5] := 0.08694311;
      W_g[6,6] := 0.12037072;
      W_g[6,7] := -0.05689518;
      W_g[6,8] := -0.04548091;
      W_g[6,9] := -0.04116108;
      W_g[6,10] := -0.11022148;
      W_g[6,11] := -0.00768893;
      W_g[6,12] := -0.00966344;
      W_g[6,13] := 0.02458816;
      W_g[6,14] := -0.01190010;
      W_g[6,15] := 0.01383197;
      W_g[6,16] := -0.06608868;
      W_g[6,17] := -0.09631553;
      W_g[6,18] := 0.00410174;
      W_g[6,19] := -0.01705389;
      W_g[6,20] := -0.12000423;
      W_g[6,21] := 0.02343578;
      W_g[6,22] := 0.01301972;
      W_g[6,23] := -0.01314613;
      W_g[6,24] := 0.03210555;
      W_g[6,25] := 0.08340400;
      W_g[6,26] := 0.00381628;
      W_g[6,27] := 0.02066490;
      W_g[6,28] := 0.13545376;
      W_g[6,29] := -0.02235859;
      W_g[6,30] := 0.00567887;
      W_g[6,31] := -0.01609200;
      W_g[6,32] := 0.00275211;
      W_g[6,33] := -0.00319188;
      W_g[6,34] := 0.29818228;
      W_g[6,35] := -0.14841233;
      W_g[6,36] := -0.03300164;
      W_g[6,37] := 0.11441298;
      W_g[6,38] := -0.02922709;
      W_g[6,39] := -0.01992949;
      W_g[7,0] := 0.00839877;
      W_g[7,1] := 0.02150501;
      W_g[7,2] := 0.01506129;
      W_g[7,3] := -0.01818663;
      W_g[7,4] := -0.00172730;
      W_g[7,5] := 0.01742283;
      W_g[7,6] := -0.02156242;
      W_g[7,7] := -0.01181841;
      W_g[7,8] := -0.01749515;
      W_g[7,9] := -0.02590540;
      W_g[7,10] := 0.00439977;
      W_g[7,11] := -0.07244217;
      W_g[7,12] := -0.06153556;
      W_g[7,13] := 0.05554190;
      W_g[7,14] := -0.08222511;
      W_g[7,15] := -0.08914689;
      W_g[7,16] := 0.00833936;
      W_g[7,17] := 0.11001267;
      W_g[7,18] := -0.03441850;
      W_g[7,19] := -0.04929563;
      W_g[7,20] := 0.01391720;
      W_g[7,21] := -0.05856322;
      W_g[7,22] := -0.00836417;
      W_g[7,23] := 0.04760852;
      W_g[7,24] := -0.36479574;
      W_g[7,25] := 0.03032077;
      W_g[7,26] := 0.04377243;
      W_g[7,27] := -0.06456570;
      W_g[7,28] := -0.00286705;
      W_g[7,29] := -0.04210155;
      W_g[7,30] := -0.01276377;
      W_g[7,31] := -0.00248455;
      W_g[7,32] := -0.01693913;
      W_g[7,33] := -0.00395950;
      W_g[7,34] := 0.09809387;
      W_g[7,35] := -0.11791219;
      W_g[7,36] := -0.04663706;
      W_g[7,37] := 0.06912785;
      W_g[7,38] := -0.04792204;
      W_g[7,39] := -0.29780853;
      W_o[0,0] := -0.24878871;
      W_o[0,1] := -0.45281693;
      W_o[0,2] := -0.05303451;
      W_o[0,3] := -0.08851492;
      W_o[0,4] := 0.39578766;
      W_o[0,5] := 0.02682471;
      W_o[0,6] := 0.23473206;
      W_o[0,7] := 0.16451281;
      W_o[0,8] := 0.06450332;
      W_o[0,9] := 0.10670687;
      W_o[0,10] := -0.07381078;
      W_o[0,11] := -0.08583919;
      W_o[0,12] := 0.10715991;
      W_o[0,13] := -0.47128552;
      W_o[0,14] := 0.22714868;
      W_o[0,15] := -0.50816250;
      W_o[0,16] := -0.11266220;
      W_o[0,17] := 0.33043900;
      W_o[0,18] := 0.49529704;
      W_o[0,19] := 0.06039276;
      W_o[0,20] := 0.15377070;
      W_o[0,21] := -0.19991648;
      W_o[0,22] := 1.07608783;
      W_o[0,23] := -0.23781183;
      W_o[0,24] := 1.15331578;
      W_o[0,25] := 1.45630133;
      W_o[0,26] := -0.30574724;
      W_o[0,27] := -0.43502858;
      W_o[0,28] := 0.13444777;
      W_o[0,29] := -0.48089328;
      W_o[0,30] := 0.87106293;
      W_o[0,31] := 0.62270272;
      W_o[0,32] := 0.42734545;
      W_o[0,33] := 0.16070290;
      W_o[0,34] := 1.78311431;
      W_o[0,35] := 0.05535344;
      W_o[0,36] := 0.18587643;
      W_o[0,37] := 0.08107077;
      W_o[0,38] := 0.27057359;
      W_o[0,39] := -0.04014807;
      W_o[1,0] := 0.17987324;
      W_o[1,1] := -0.20177005;
      W_o[1,2] := -0.23272584;
      W_o[1,3] := -0.06171975;
      W_o[1,4] := 0.16163252;
      W_o[1,5] := 0.04768089;
      W_o[1,6] := -0.01735293;
      W_o[1,7] := -0.00856016;
      W_o[1,8] := 0.32226062;
      W_o[1,9] := 0.14564918;
      W_o[1,10] := 0.34103507;
      W_o[1,11] := -0.47851020;
      W_o[1,12] := -0.16536747;
      W_o[1,13] := -0.07199546;
      W_o[1,14] := 0.38576946;
      W_o[1,15] := 0.15553798;
      W_o[1,16] := 0.16951348;
      W_o[1,17] := -0.34140691;
      W_o[1,18] := 0.54336584;
      W_o[1,19] := -0.39412004;
      W_o[1,20] := -0.18107198;
      W_o[1,21] := 0.08229911;
      W_o[1,22] := 0.34285191;
      W_o[1,23] := -0.38594139;
      W_o[1,24] := 1.56069613;
      W_o[1,25] := 1.31107664;
      W_o[1,26] := -0.07977130;
      W_o[1,27] := -0.00066841;
      W_o[1,28] := 0.02706419;
      W_o[1,29] := -0.53140843;
      W_o[1,30] := 0.82663709;
      W_o[1,31] := 0.20585302;
      W_o[1,32] := 0.26289618;
      W_o[1,33] := 0.05673197;
      W_o[1,34] := 1.33109844;
      W_o[1,35] := 0.65518051;
      W_o[1,36] := -0.04780313;
      W_o[1,37] := 0.11147591;
      W_o[1,38] := 0.46894863;
      W_o[1,39] := 0.01827455;
      W_o[2,0] := -0.13741741;
      W_o[2,1] := 0.34161562;
      W_o[2,2] := 0.00265318;
      W_o[2,3] := -0.06815082;
      W_o[2,4] := -0.63534689;
      W_o[2,5] := 0.09096143;
      W_o[2,6] := 0.18871199;
      W_o[2,7] := -0.03421344;
      W_o[2,8] := -0.00024948;
      W_o[2,9] := -0.13563773;
      W_o[2,10] := 0.15499417;
      W_o[2,11] := 0.10373094;
      W_o[2,12] := -0.09785850;
      W_o[2,13] := 0.08585915;
      W_o[2,14] := 0.04649240;
      W_o[2,15] := 0.01026138;
      W_o[2,16] := -0.04262185;
      W_o[2,17] := -0.01874319;
      W_o[2,18] := 0.75688982;
      W_o[2,19] := -0.04560044;
      W_o[2,20] := -0.32223263;
      W_o[2,21] := 0.10837347;
      W_o[2,22] := 0.36421233;
      W_o[2,23] := 0.10329347;
      W_o[2,24] := -0.27218717;
      W_o[2,25] := 0.17619081;
      W_o[2,26] := -0.18144348;
      W_o[2,27] := -0.17446589;
      W_o[2,28] := 0.09568179;
      W_o[2,29] := 0.39024752;
      W_o[2,30] := 0.31926751;
      W_o[2,31] := -0.09343637;
      W_o[2,32] := -0.04776040;
      W_o[2,33] := -0.04253375;
      W_o[2,34] := -0.02549809;
      W_o[2,35] := 0.12155074;
      W_o[2,36] := -0.12728153;
      W_o[2,37] := -0.06793334;
      W_o[2,38] := 0.03087276;
      W_o[2,39] := 0.05013068;
      W_o[3,0] := -0.15653051;
      W_o[3,1] := -0.04078253;
      W_o[3,2] := -0.21346539;
      W_o[3,3] := -0.16302916;
      W_o[3,4] := -0.13266797;
      W_o[3,5] := -0.05849253;
      W_o[3,6] := 0.00807450;
      W_o[3,7] := 0.08821388;
      W_o[3,8] := 0.15438399;
      W_o[3,9] := -0.24945748;
      W_o[3,10] := 0.03148121;
      W_o[3,11] := 0.17463362;
      W_o[3,12] := -0.24076079;
      W_o[3,13] := -0.05835954;
      W_o[3,14] := 0.00083490;
      W_o[3,15] := -0.05821047;
      W_o[3,16] := 0.22283494;
      W_o[3,17] := 0.27039650;
      W_o[3,18] := 0.03926261;
      W_o[3,19] := 0.13555294;
      W_o[3,20] := 0.25270861;
      W_o[3,21] := 0.50729799;
      W_o[3,22] := -0.15098204;
      W_o[3,23] := -0.02635484;
      W_o[3,24] := -0.16301835;
      W_o[3,25] := 0.03315194;
      W_o[3,26] := 0.17386480;
      W_o[3,27] := -0.04533337;
      W_o[3,28] := -0.26984090;
      W_o[3,29] := 0.12042534;
      W_o[3,30] := -0.05481909;
      W_o[3,31] := -0.07778496;
      W_o[3,32] := -0.12814386;
      W_o[3,33] := 0.41067052;
      W_o[3,34] := -0.04621636;
      W_o[3,35] := -0.08714477;
      W_o[3,36] := -0.20655701;
      W_o[3,37] := -0.03565258;
      W_o[3,38] := -0.08211713;
      W_o[3,39] := -0.11460824;
      W_o[4,0] := -0.16526031;
      W_o[4,1] := -0.03820162;
      W_o[4,2] := 0.23743653;
      W_o[4,3] := -0.17364512;
      W_o[4,4] := 0.09611007;
      W_o[4,5] := 0.25984883;
      W_o[4,6] := 0.24360292;
      W_o[4,7] := 0.08559894;
      W_o[4,8] := -0.02284659;
      W_o[4,9] := 0.20195185;
      W_o[4,10] := -0.09046014;
      W_o[4,11] := 0.09581435;
      W_o[4,12] := -0.15597157;
      W_o[4,13] := -0.34664866;
      W_o[4,14] := 0.11788706;
      W_o[4,15] := 0.03617490;
      W_o[4,16] := -0.19772679;
      W_o[4,17] := -0.27061427;
      W_o[4,18] := -0.07025576;
      W_o[4,19] := -0.20179892;
      W_o[4,20] := -0.13330138;
      W_o[4,21] := 0.28108272;
      W_o[4,22] := -0.04382841;
      W_o[4,23] := -0.38677481;
      W_o[4,24] := -0.51250386;
      W_o[4,25] := -0.38813958;
      W_o[4,26] := -0.04432906;
      W_o[4,27] := -0.18282278;
      W_o[4,28] := 0.06468461;
      W_o[4,29] := -0.34807864;
      W_o[4,30] := -0.41589615;
      W_o[4,31] := 0.16075355;
      W_o[4,32] := 0.15460733;
      W_o[4,33] := 0.22832997;
      W_o[4,34] := 0.03074585;
      W_o[4,35] := 0.02588873;
      W_o[4,36] := -0.19890888;
      W_o[4,37] := 0.17934620;
      W_o[4,38] := -0.07465497;
      W_o[4,39] := 0.18535613;
      W_o[5,0] := 0.35529122;
      W_o[5,1] := -0.45068535;
      W_o[5,2] := 0.13398276;
      W_o[5,3] := 0.00250324;
      W_o[5,4] := 0.09135553;
      W_o[5,5] := 0.33329329;
      W_o[5,6] := -0.15334524;
      W_o[5,7] := 0.03885195;
      W_o[5,8] := -0.61340588;
      W_o[5,9] := -0.08592401;
      W_o[5,10] := -0.11830733;
      W_o[5,11] := -0.17615788;
      W_o[5,12] := -0.24301590;
      W_o[5,13] := -0.17049399;
      W_o[5,14] := 0.19884115;
      W_o[5,15] := -0.07459871;
      W_o[5,16] := -0.47671059;
      W_o[5,17] := 0.14353496;
      W_o[5,18] := 0.69755995;
      W_o[5,19] := -0.29544228;
      W_o[5,20] := -0.03883540;
      W_o[5,21] := -0.22129694;
      W_o[5,22] := 0.11786394;
      W_o[5,23] := -0.10525186;
      W_o[5,24] := 1.27088118;
      W_o[5,25] := 1.08401871;
      W_o[5,26] := -0.37344339;
      W_o[5,27] := -0.23756148;
      W_o[5,28] := 0.06141074;
      W_o[5,29] := 0.13355421;
      W_o[5,30] := 0.34222761;
      W_o[5,31] := -0.05769080;
      W_o[5,32] := 0.44572812;
      W_o[5,33] := -0.13044961;
      W_o[5,34] := 0.44415033;
      W_o[5,35] := -0.15364335;
      W_o[5,36] := -0.08437125;
      W_o[5,37] := -0.08841761;
      W_o[5,38] := 0.11458829;
      W_o[5,39] := 0.62695736;
      W_o[6,0] := 0.03065801;
      W_o[6,1] := 0.03260401;
      W_o[6,2] := -0.19908448;
      W_o[6,3] := 0.10675497;
      W_o[6,4] := -0.02801576;
      W_o[6,5] := 0.32186738;
      W_o[6,6] := 1.07099915;
      W_o[6,7] := -0.22513410;
      W_o[6,8] := 0.08130264;
      W_o[6,9] := -0.11853161;
      W_o[6,10] := 0.28825247;
      W_o[6,11] := -0.34321690;
      W_o[6,12] := 0.40200213;
      W_o[6,13] := -0.02302332;
      W_o[6,14] := 0.01709228;
      W_o[6,15] := -0.03287499;
      W_o[6,16] := 0.35959429;
      W_o[6,17] := 0.28991431;
      W_o[6,18] := 0.26372039;
      W_o[6,19] := -0.17363600;
      W_o[6,20] := -0.96958780;
      W_o[6,21] := 0.27258980;
      W_o[6,22] := 1.01800835;
      W_o[6,23] := -0.45700833;
      W_o[6,24] := 1.27344668;
      W_o[6,25] := 0.80010319;
      W_o[6,26] := 0.50079250;
      W_o[6,27] := -0.00981760;
      W_o[6,28] := 0.39598280;
      W_o[6,29] := -0.44397491;
      W_o[6,30] := 1.02373374;
      W_o[6,31] := -0.20951441;
      W_o[6,32] := 0.59132648;
      W_o[6,33] := -0.03599635;
      W_o[6,34] := 1.37534094;
      W_o[6,35] := 0.25570524;
      W_o[6,36] := 0.01851447;
      W_o[6,37] := 0.41994217;
      W_o[6,38] := -0.12552960;
      W_o[6,39] := 0.69572401;
      W_o[7,0] := -0.21226366;
      W_o[7,1] := -0.04577332;
      W_o[7,2] := 0.12693021;
      W_o[7,3] := -0.00553917;
      W_o[7,4] := 0.31903967;
      W_o[7,5] := 0.28985706;
      W_o[7,6] := 0.07334051;
      W_o[7,7] := 0.07537151;
      W_o[7,8] := -0.06602987;
      W_o[7,9] := 0.10063405;
      W_o[7,10] := -0.07167389;
      W_o[7,11] := -0.64208913;
      W_o[7,12] := 0.26317602;
      W_o[7,13] := -0.19404016;
      W_o[7,14] := -0.57089996;
      W_o[7,15] := -0.06107605;
      W_o[7,16] := 0.04890145;
      W_o[7,17] := 0.32024038;
      W_o[7,18] := 0.51453072;
      W_o[7,19] := -0.12590186;
      W_o[7,20] := 0.02570236;
      W_o[7,21] := 0.33773011;
      W_o[7,22] := 0.03015064;
      W_o[7,23] := -0.46817833;
      W_o[7,24] := 1.17787540;
      W_o[7,25] := 1.11605489;
      W_o[7,26] := -0.33396244;
      W_o[7,27] := -0.07750119;
      W_o[7,28] := -0.24094582;
      W_o[7,29] := -0.19267891;
      W_o[7,30] := 0.28351098;
      W_o[7,31] := 0.11068187;
      W_o[7,32] := -0.11161529;
      W_o[7,33] := 0.05576994;
      W_o[7,34] := 0.15852658;
      W_o[7,35] := 0.19595769;
      W_o[7,36] := 0.17078656;
      W_o[7,37] := 0.12906086;
      W_o[7,38] := 0.20672542;
      W_o[7,39] := 0.13961391;
      R_i[0,0] := -0.29720330;
      R_i[0,1] := -0.05501601;
      R_i[0,2] := 0.19428261;
      R_i[0,3] := -0.01147678;
      R_i[0,4] := -0.35804778;
      R_i[0,5] := 0.35627866;
      R_i[0,6] := 0.06648605;
      R_i[0,7] := -0.25248384;
      R_i[1,0] := -0.00485134;
      R_i[1,1] := 0.29569951;
      R_i[1,2] := 0.46215025;
      R_i[1,3] := -0.32642034;
      R_i[1,4] := 0.30512771;
      R_i[1,5] := -0.08773772;
      R_i[1,6] := -0.13170604;
      R_i[1,7] := 0.15243977;
      R_i[2,0] := 0.20030405;
      R_i[2,1] := 0.22486736;
      R_i[2,2] := -0.26627916;
      R_i[2,3] := 0.21764944;
      R_i[2,4] := -0.39947459;
      R_i[2,5] := 0.41491815;
      R_i[2,6] := 0.27285352;
      R_i[2,7] := 0.31419027;
      R_i[3,0] := 0.15271637;
      R_i[3,1] := 0.13401978;
      R_i[3,2] := -0.02607298;
      R_i[3,3] := -0.29988387;
      R_i[3,4] := -0.16316661;
      R_i[3,5] := 0.33023968;
      R_i[3,6] := 0.17649920;
      R_i[3,7] := 0.19594158;
      R_i[4,0] := 0.24785545;
      R_i[4,1] := 0.03621851;
      R_i[4,2] := 0.76205403;
      R_i[4,3] := -0.31073129;
      R_i[4,4] := -0.09589436;
      R_i[4,5] := 0.18456733;
      R_i[4,6] := -0.57247859;
      R_i[4,7] := -0.15726174;
      R_i[5,0] := -0.15299343;
      R_i[5,1] := 0.06710675;
      R_i[5,2] := 0.64831352;
      R_i[5,3] := -0.22750993;
      R_i[5,4] := -0.76823664;
      R_i[5,5] := 0.37383676;
      R_i[5,6] := 0.17858171;
      R_i[5,7] := 0.35545036;
      R_i[6,0] := -0.04436296;
      R_i[6,1] := 0.33972314;
      R_i[6,2] := 0.23785813;
      R_i[6,3] := 0.20984678;
      R_i[6,4] := -0.05630715;
      R_i[6,5] := 0.25487366;
      R_i[6,6] := -0.22129624;
      R_i[6,7] := -0.10079595;
      R_i[7,0] := 0.19636191;
      R_i[7,1] := 0.40730953;
      R_i[7,2] := 0.74057549;
      R_i[7,3] := 0.11769681;
      R_i[7,4] := -0.07874840;
      R_i[7,5] := 0.13999742;
      R_i[7,6] := -0.07538932;
      R_i[7,7] := 0.15130904;
      R_f[0,0] := -0.15415196;
      R_f[0,1] := 0.14001700;
      R_f[0,2] := 0.32896742;
      R_f[0,3] := 0.03486477;
      R_f[0,4] := -0.25475094;
      R_f[0,5] := 0.25555649;
      R_f[0,6] := 0.16113877;
      R_f[0,7] := -0.19586459;
      R_f[1,0] := 0.28900579;
      R_f[1,1] := 0.51801419;
      R_f[1,2] := 0.41163966;
      R_f[1,3] := -0.49210873;
      R_f[1,4] := -0.44169796;
      R_f[1,5] := 0.52491426;
      R_f[1,6] := 0.09079631;
      R_f[1,7] := 0.24646547;
      R_f[2,0] := 0.33840427;
      R_f[2,1] := 0.31135768;
      R_f[2,2] := -0.55702937;
      R_f[2,3] := -0.14924698;
      R_f[2,4] := 0.16647284;
      R_f[2,5] := -0.04085749;
      R_f[2,6] := -0.02604689;
      R_f[2,7] := -0.17268968;
      R_f[3,0] := 0.32577130;
      R_f[3,1] := 0.36095178;
      R_f[3,2] := 0.43605298;
      R_f[3,3] := 0.16874421;
      R_f[3,4] := -0.12284465;
      R_f[3,5] := 0.03751094;
      R_f[3,6] := 0.02462184;
      R_f[3,7] := 0.03318978;
      R_f[4,0] := 0.49182421;
      R_f[4,1] := 0.16429330;
      R_f[4,2] := 0.53267479;
      R_f[4,3] := -0.49470288;
      R_f[4,4] := 0.10341619;
      R_f[4,5] := -0.07133373;
      R_f[4,6] := 0.11399978;
      R_f[4,7] := -0.19527824;
      R_f[5,0] := 0.27028599;
      R_f[5,1] := 0.05122235;
      R_f[5,2] := -0.27298668;
      R_f[5,3] := 0.00193437;
      R_f[5,4] := -0.21285854;
      R_f[5,5] := 0.08526506;
      R_f[5,6] := -0.23500830;
      R_f[5,7] := 0.12631051;
      R_f[6,0] := 0.71271533;
      R_f[6,1] := 0.45810968;
      R_f[6,2] := 0.05682573;
      R_f[6,3] := -0.70776463;
      R_f[6,4] := -0.22887982;
      R_f[6,5] := 0.43033603;
      R_f[6,6] := -0.06712849;
      R_f[6,7] := -0.50418854;
      R_f[7,0] := -0.08720636;
      R_f[7,1] := 0.07314771;
      R_f[7,2] := -0.10617252;
      R_f[7,3] := -0.22731772;
      R_f[7,4] := -0.38440135;
      R_f[7,5] := 0.22375256;
      R_f[7,6] := 0.19357640;
      R_f[7,7] := 0.02181435;
      R_g[0,0] := -1.67002046;
      R_g[0,1] := 0.22261654;
      R_g[0,2] := -0.29516104;
      R_g[0,3] := 0.38097781;
      R_g[0,4] := 0.18069918;
      R_g[0,5] := -0.04807178;
      R_g[0,6] := -0.21403493;
      R_g[0,7] := 0.30647677;
      R_g[1,0] := 0.09286369;
      R_g[1,1] := -1.67246938;
      R_g[1,2] := 0.25422445;
      R_g[1,3] := -0.13823049;
      R_g[1,4] := -0.05546627;
      R_g[1,5] := 0.02552741;
      R_g[1,6] := -0.04196908;
      R_g[1,7] := -0.12302180;
      R_g[2,0] := 0.12508599;
      R_g[2,1] := -0.01198944;
      R_g[2,2] := -1.76017654;
      R_g[2,3] := 0.41029209;
      R_g[2,4] := 0.32856131;
      R_g[2,5] := 0.19418783;
      R_g[2,6] := 0.13047464;
      R_g[2,7] := 0.06735183;
      R_g[3,0] := -0.08110875;
      R_g[3,1] := 0.12964080;
      R_g[3,2] := 0.03910316;
      R_g[3,3] := -1.58626795;
      R_g[3,4] := 0.05309961;
      R_g[3,5] := 0.19302739;
      R_g[3,6] := -0.03232419;
      R_g[3,7] := 0.10759025;
      R_g[4,0] := 0.10843568;
      R_g[4,1] := -0.08969119;
      R_g[4,2] := 0.47807658;
      R_g[4,3] := -0.48509952;
      R_g[4,4] := -1.74958336;
      R_g[4,5] := -0.07144331;
      R_g[4,6] := -0.06208268;
      R_g[4,7] := -0.12589887;
      R_g[5,0] := -0.01311982;
      R_g[5,1] := -0.07684252;
      R_g[5,2] := 0.20680495;
      R_g[5,3] := -0.38980842;
      R_g[5,4] := -0.04986978;
      R_g[5,5] := -1.06202638;
      R_g[5,6] := 0.11428019;
      R_g[5,7] := -0.20394331;
      R_g[6,0] := 0.06553666;
      R_g[6,1] := -0.05139922;
      R_g[6,2] := 0.44536793;
      R_g[6,3] := -0.27498397;
      R_g[6,4] := -0.32525745;
      R_g[6,5] := 0.00937504;
      R_g[6,6] := -1.56192875;
      R_g[6,7] := -0.11409894;
      R_g[7,0] := 0.05325243;
      R_g[7,1] := -0.33739990;
      R_g[7,2] := 0.21331263;
      R_g[7,3] := -0.37539151;
      R_g[7,4] := -0.17099947;
      R_g[7,5] := 0.00843642;
      R_g[7,6] := 0.11368373;
      R_g[7,7] := -1.43479502;
      R_o[0,0] := 0.28625217;
      R_o[0,1] := 0.62617600;
      R_o[0,2] := 0.51247001;
      R_o[0,3] := -0.33488548;
      R_o[0,4] := -0.78386301;
      R_o[0,5] := 0.73291373;
      R_o[0,6] := -1.09786367;
      R_o[0,7] := -0.31238851;
      R_o[1,0] := 0.43348855;
      R_o[1,1] := 0.54565865;
      R_o[1,2] := 0.52155811;
      R_o[1,3] := -0.07661161;
      R_o[1,4] := -0.77065903;
      R_o[1,5] := 0.33984208;
      R_o[1,6] := -0.21829525;
      R_o[1,7] := 0.30410659;
      R_o[2,0] := 0.77740079;
      R_o[2,1] := 0.77948558;
      R_o[2,2] := 0.25081304;
      R_o[2,3] := 0.22476536;
      R_o[2,4] := -0.18188496;
      R_o[2,5] := 0.24920675;
      R_o[2,6] := -0.32646251;
      R_o[2,7] := -0.22284411;
      R_o[3,0] := 0.10846130;
      R_o[3,1] := 0.15308166;
      R_o[3,2] := 0.98173195;
      R_o[3,3] := -0.20129372;
      R_o[3,4] := -0.48236448;
      R_o[3,5] := 0.29829371;
      R_o[3,6] := -0.59647918;
      R_o[3,7] := -0.13544692;
      R_o[4,0] := 0.64042091;
      R_o[4,1] := -0.19734913;
      R_o[4,2] := 1.14491618;
      R_o[4,3] := -0.14366756;
      R_o[4,4] := -0.72905266;
      R_o[4,5] := 0.17306720;
      R_o[4,6] := 0.00839791;
      R_o[4,7] := 0.25284833;
      R_o[5,0] := 0.54454422;
      R_o[5,1] := 0.86287361;
      R_o[5,2] := 0.75096619;
      R_o[5,3] := 0.13229862;
      R_o[5,4] := -0.27491441;
      R_o[5,5] := 0.70543158;
      R_o[5,6] := -0.11946990;
      R_o[5,7] := 0.17286766;
      R_o[6,0] := 0.77812266;
      R_o[6,1] := 0.48867458;
      R_o[6,2] := 0.87114924;
      R_o[6,3] := 0.21844880;
      R_o[6,4] := -0.41514960;
      R_o[6,5] := -0.14079522;
      R_o[6,6] := -0.10740466;
      R_o[6,7] := -0.09739928;
      R_o[7,0] := 0.68203056;
      R_o[7,1] := 0.50477397;
      R_o[7,2] := 0.62449515;
      R_o[7,3] := 0.17028584;
      R_o[7,4] := -0.56497252;
      R_o[7,5] := 0.31056079;
      R_o[7,6] := -0.29031694;
      R_o[7,7] := 0.44926986;
      B_i[0] := 0.85732204;
      B_i[1] := 1.04156196;
      B_i[2] := 0.97363615;
      B_i[3] := 0.80207175;
      B_i[4] := 0.80256236;
      B_i[5] := 1.98055279;
      B_i[6] := 1.54851460;
      B_i[7] := 1.91203833;
      B_f[0] := 0.74003136;
      B_f[1] := 1.29651260;
      B_f[2] := 1.39809060;
      B_f[3] := 1.21004391;
      B_f[4] := 0.88460255;
      B_f[5] := -0.01221798;
      B_f[6] := 1.10466242;
      B_f[7] := 0.64986908;
      B_g[0] := 0.31623846;
      B_g[1] := 0.62138993;
      B_g[2] := 0.74492103;
      B_g[3] := -0.47756320;
      B_g[4] := -0.68758571;
      B_g[5] := 0.16762234;
      B_g[6] := -0.50441682;
      B_g[7] := -0.09181471;
      B_o[0] := 3.19267225;
      B_o[1] := 2.76363182;
      B_o[2] := 2.40052104;
      B_o[3] := 2.11938143;
      B_o[4] := 2.60010386;
      B_o[5] := 2.18173027;
      B_o[6] := 2.06268406;
      B_o[7] := 2.10852313;
      FC_W[0,0] := -0.79911309;
      FC_W[0,1] := -0.93833846;
      FC_W[0,2] := 1.09520888;
      FC_W[0,3] := 0.43509555;
      FC_W[0,4] := -0.35498026;
      FC_W[0,5] := 1.23117495;
      FC_W[0,6] := 0.54596531;
      FC_W[0,7] := -0.04457461;
      FC_W[1,0] := 0.30732417;
      FC_W[1,1] := 0.80071634;
      FC_W[1,2] := 0.71018058;
      FC_W[1,3] := -0.61475515;
      FC_W[1,4] := -1.05773103;
      FC_W[1,5] := -1.65802586;
      FC_W[1,6] := -0.15574944;
      FC_W[1,7] := 0.56488359;
      FC_W[2,0] := -0.79928327;
      FC_W[2,1] := -0.89827907;
      FC_W[2,2] := 1.07494175;
      FC_W[2,3] := 0.43071118;
      FC_W[2,4] := -0.31526205;
      FC_W[2,5] := 1.24351621;
      FC_W[2,6] := 0.53584868;
      FC_W[2,7] := -0.07105654;
      FC_W[3,0] := 0.06145537;
      FC_W[3,1] := -0.07917563;
      FC_W[3,2] := 0.47143328;
      FC_W[3,3] := -0.97099501;
      FC_W[3,4] := 0.77169645;
      FC_W[3,5] := 1.17534721;
      FC_W[3,6] := -0.98506945;
      FC_W[3,7] := -0.68494749;
      FC_W[4,0] := -1.87392640;
      FC_W[4,1] := -0.71319950;
      FC_W[4,2] := -0.97656369;
      FC_W[4,3] := -1.93710411;
      FC_W[4,4] := -0.74523616;
      FC_W[4,5] := 0.40530244;
      FC_W[4,6] := 0.01008961;
      FC_W[4,7] := -0.04781210;
      FC_W[5,0] := 0.22815995;
      FC_W[5,1] := 0.40298557;
      FC_W[5,2] := 0.48270676;
      FC_W[5,3] := -0.44884250;
      FC_W[5,4] := 0.74876332;
      FC_W[5,5] := -0.57336783;
      FC_W[5,6] := 1.27662027;
      FC_W[5,7] := 0.50955653;
      FC_W[6,0] := 1.13151014;
      FC_W[6,1] := -0.50774103;
      FC_W[6,2] := 0.43078673;
      FC_W[6,3] := -1.29680264;
      FC_W[6,4] := 1.18923640;
      FC_W[6,5] := 0.02214067;
      FC_W[6,6] := 1.83503294;
      FC_W[6,7] := -0.65552771;
      FC_W[7,0] := 0.06186135;
      FC_W[7,1] := -0.09877446;
      FC_W[7,2] := 0.47054976;
      FC_W[7,3] := -0.97938317;
      FC_W[7,4] := 0.76673663;
      FC_W[7,5] := 1.18406940;
      FC_W[7,6] := -0.97699875;
      FC_W[7,7] := -0.68285751;
      FC_W[8,0] := 0.05534381;
      FC_W[8,1] := -0.06393234;
      FC_W[8,2] := 0.42852098;
      FC_W[8,3] := -0.91158271;
      FC_W[8,4] := 0.81992948;
      FC_W[8,5] := 1.17474234;
      FC_W[8,6] := -0.96696079;
      FC_W[8,7] := -0.64814442;
      FC_W[9,0] := 0.06112890;
      FC_W[9,1] := -0.08640661;
      FC_W[9,2] := 0.48090583;
      FC_W[9,3] := -0.96519989;
      FC_W[9,4] := 0.76665956;
      FC_W[9,5] := 1.17957020;
      FC_W[9,6] := -0.98317134;
      FC_W[9,7] := -0.67911482;
      FC_W[10,0] := -0.55945873;
      FC_W[10,1] := 0.50921994;
      FC_W[10,2] := 0.39391521;
      FC_W[10,3] := -0.05040882;
      FC_W[10,4] := 0.13381737;
      FC_W[10,5] := 0.80598813;
      FC_W[10,6] := -1.79597354;
      FC_W[10,7] := 0.09913790;
      FC_W[11,0] := 0.09679934;
      FC_W[11,1] := 1.45000255;
      FC_W[11,2] := -0.34398675;
      FC_W[11,3] := -0.65334404;
      FC_W[11,4] := -0.48840344;
      FC_W[11,5] := 0.45034793;
      FC_W[11,6] := 0.20451836;
      FC_W[11,7] := -1.16122139;
      FC_W[12,0] := 0.31311855;
      FC_W[12,1] := 1.34233701;
      FC_W[12,2] := -0.30392364;
      FC_W[12,3] := -0.89511561;
      FC_W[12,4] := -0.31252480;
      FC_W[12,5] := 0.42357349;
      FC_W[12,6] := -0.04789438;
      FC_W[12,7] := -0.95470685;
      FC_W[13,0] := -0.67863357;
      FC_W[13,1] := 0.55870867;
      FC_W[13,2] := 2.74645376;
      FC_W[13,3] := -0.54551154;
      FC_W[13,4] := -1.40819108;
      FC_W[13,5] := -0.65208882;
      FC_W[13,6] := -0.04722747;
      FC_W[13,7] := 1.13449383;
      FC_W[14,0] := -1.63870704;
      FC_W[14,1] := -1.43244660;
      FC_W[14,2] := 1.88617778;
      FC_W[14,3] := -0.14083456;
      FC_W[14,4] := 1.25434613;
      FC_W[14,5] := -1.56908119;
      FC_W[14,6] := -0.79074830;
      FC_W[14,7] := -2.52818203;
      FC_W[15,0] := -0.22405152;
      FC_W[15,1] := 1.40958560;
      FC_W[15,2] := -0.12493899;
      FC_W[15,3] := -0.39721119;
      FC_W[15,4] := -0.52675790;
      FC_W[15,5] := 0.29834321;
      FC_W[15,6] := 0.42443123;
      FC_W[15,7] := -1.51365042;
      FC_W[16,0] := -0.35442686;
      FC_W[16,1] := -1.87087142;
      FC_W[16,2] := 1.28207767;
      FC_W[16,3] := -1.00388706;
      FC_W[16,4] := 1.52664959;
      FC_W[16,5] := -0.90419412;
      FC_W[16,6] := -1.65340745;
      FC_W[16,7] := -0.85398114;
      FC_W[17,0] := 1.81199193;
      FC_W[17,1] := -0.77926898;
      FC_W[17,2] := -0.48014465;
      FC_W[17,3] := -1.65164447;
      FC_W[17,4] := 1.07409704;
      FC_W[17,5] := 0.35728425;
      FC_W[17,6] := -1.67923045;
      FC_W[17,7] := 2.20978189;
      FC_W[18,0] := 0.59539229;
      FC_W[18,1] := -1.52473056;
      FC_W[18,2] := -1.85000372;
      FC_W[18,3] := -0.20748819;
      FC_W[18,4] := -0.57798457;
      FC_W[18,5] := 0.85016835;
      FC_W[18,6] := 0.29200807;
      FC_W[18,7] := -1.38809645;
      FC_W[19,0] := 0.19826975;
      FC_W[19,1] := 1.70039785;
      FC_W[19,2] := 0.07619762;
      FC_W[19,3] := -0.80908722;
      FC_W[19,4] := -0.19027834;
      FC_W[19,5] := 0.20950752;
      FC_W[19,6] := -0.03333457;
      FC_W[19,7] := -0.61634111;
      FC_W[20,0] := -1.09664285;
      FC_W[20,1] := 0.29726404;
      FC_W[20,2] := -0.01492481;
      FC_W[20,3] := 0.46071255;
      FC_W[20,4] := -1.59879112;
      FC_W[20,5] := 0.02794913;
      FC_W[20,6] := -1.93254459;
      FC_W[20,7] := 0.38252020;
      FC_W[21,0] := 2.34788537;
      FC_W[21,1] := -1.36648786;
      FC_W[21,2] := 0.24216530;
      FC_W[21,3] := -0.22190996;
      FC_W[21,4] := -0.50946277;
      FC_W[21,5] := 0.37187195;
      FC_W[21,6] := 0.68050140;
      FC_W[21,7] := -1.89826512;
      FC_W[22,0] := 0.34295273;
      FC_W[22,1] := -0.70024264;
      FC_W[22,2] := 2.52141047;
      FC_W[22,3] := -2.68626642;
      FC_W[22,4] := -2.60129905;
      FC_W[22,5] := -0.34002843;
      FC_W[22,6] := -0.65852845;
      FC_W[22,7] := -0.88338953;
      FC_W[23,0] := -0.82124501;
      FC_W[23,1] := 0.75074446;
      FC_W[23,2] := 2.99681067;
      FC_W[23,3] := -0.67825657;
      FC_W[23,4] := -0.94996166;
      FC_W[23,5] := -0.26541135;
      FC_W[23,6] := -0.71499181;
      FC_W[23,7] := 0.85002565;
      FC_W[24,0] := 0.39461923;
      FC_W[24,1] := -0.77516311;
      FC_W[24,2] := 2.46279955;
      FC_W[24,3] := -2.73454237;
      FC_W[24,4] := -2.63833332;
      FC_W[24,5] := -0.31525555;
      FC_W[24,6] := -0.61657113;
      FC_W[24,7] := -0.96707428;
      FC_W[25,0] := 0.39434937;
      FC_W[25,1] := -0.77477384;
      FC_W[25,2] := 2.46124387;
      FC_W[25,3] := -2.73295689;
      FC_W[25,4] := -2.63696575;
      FC_W[25,5] := -0.31505886;
      FC_W[25,6] := -0.61616051;
      FC_W[25,7] := -0.96655226;
      FC_W[26,0] := -1.25524557;
      FC_W[26,1] := 0.68099910;
      FC_W[26,2] := 2.24707365;
      FC_W[26,3] := -1.90008891;
      FC_W[26,4] := -1.23129189;
      FC_W[26,5] := -0.68385196;
      FC_W[26,6] := -0.70202827;
      FC_W[26,7] := 0.85420585;
      FC_W[27,0] := 2.20356202;
      FC_W[27,1] := -1.34705377;
      FC_W[27,2] := -0.24984661;
      FC_W[27,3] := 0.19494583;
      FC_W[27,4] := -0.27059293;
      FC_W[27,5] := 0.49716923;
      FC_W[27,6] := 0.68631184;
      FC_W[27,7] := -1.82476807;
      FC_W[28,0] := -1.46181500;
      FC_W[28,1] := -0.34316191;
      FC_W[28,2] := -0.46657822;
      FC_W[28,3] := -2.00234008;
      FC_W[28,4] := 0.44393504;
      FC_W[28,5] := 0.32037762;
      FC_W[28,6] := 1.59235418;
      FC_W[28,7] := 0.08116318;
      FC_W[29,0] := -0.41624770;
      FC_W[29,1] := 0.67810297;
      FC_W[29,2] := -2.39604473;
      FC_W[29,3] := 2.50969100;
      FC_W[29,4] := 2.43244958;
      FC_W[29,5] := 0.34069127;
      FC_W[29,6] := 0.63509458;
      FC_W[29,7] := 0.85426724;
      FC_W[30,0] := 0.33883870;
      FC_W[30,1] := -0.69733250;
      FC_W[30,2] := 2.52243900;
      FC_W[30,3] := -2.68499517;
      FC_W[30,4] := -2.60072398;
      FC_W[30,5] := -0.34062445;
      FC_W[30,6] := -0.66011596;
      FC_W[30,7] := -0.87961990;
      FC_W[31,0] := 0.31169829;
      FC_W[31,1] := -0.67098248;
      FC_W[31,2] := 2.52186966;
      FC_W[31,3] := -2.67077470;
      FC_W[31,4] := -2.55351281;
      FC_W[31,5] := -0.34580857;
      FC_W[31,6] := -0.66304654;
      FC_W[31,7] := -0.84584129;
      FC_W[32,0] := 0.42391488;
      FC_W[32,1] := -0.77404338;
      FC_W[32,2] := 2.48852396;
      FC_W[32,3] := -2.73408318;
      FC_W[32,4] := -2.63075829;
      FC_W[32,5] := -0.32349947;
      FC_W[32,6] := -0.60429329;
      FC_W[32,7] := -0.96998984;
      FC_W[33,0] := 0.42112416;
      FC_W[33,1] := -0.74305284;
      FC_W[33,2] := 2.48353839;
      FC_W[33,3] := -2.72027206;
      FC_W[33,4] := -2.57575727;
      FC_W[33,5] := -0.34379905;
      FC_W[33,6] := -0.60176629;
      FC_W[33,7] := -0.93384212;
      FC_W[34,0] := 0.38578042;
      FC_W[34,1] := -0.73361003;
      FC_W[34,2] := 2.49397111;
      FC_W[34,3] := -2.70783997;
      FC_W[34,4] := -2.58508277;
      FC_W[34,5] := -0.33692864;
      FC_W[34,6] := -0.62745452;
      FC_W[34,7] := -0.91552860;
      FC_W[35,0] := 0.44358394;
      FC_W[35,1] := -0.80064774;
      FC_W[35,2] := 2.47607827;
      FC_W[35,3] := -2.71811557;
      FC_W[35,4] := -2.64654303;
      FC_W[35,5] := -0.30309862;
      FC_W[35,6] := -0.58877528;
      FC_W[35,7] := -0.99631965;
      FC_W[36,0] := 1.03216982;
      FC_W[36,1] := -1.31236815;
      FC_W[36,2] := 0.79231286;
      FC_W[36,3] := -1.15934968;
      FC_W[36,4] := -2.29796004;
      FC_W[36,5] := 0.26195404;
      FC_W[36,6] := -0.50553924;
      FC_W[36,7] := -1.66059065;
      FC_W[37,0] := 0.46099925;
      FC_W[37,1] := -0.80687803;
      FC_W[37,2] := 2.47530270;
      FC_W[37,3] := -2.70996881;
      FC_W[37,4] := -2.64459825;
      FC_W[37,5] := -0.30008873;
      FC_W[37,6] := -0.57691818;
      FC_W[37,7] := -1.00765979;
      FC_W[38,0] := -1.48978579;
      FC_W[38,1] := -1.78936589;
      FC_W[38,2] := 1.91299665;
      FC_W[38,3] := -0.32968995;
      FC_W[38,4] := 1.36646545;
      FC_W[38,5] := -1.46659601;
      FC_W[38,6] := -1.12252676;
      FC_W[38,7] := -2.30282712;
      FC_W[39,0] := -1.69402015;
      FC_W[39,1] := -1.80726838;
      FC_W[39,2] := 2.09063578;
      FC_W[39,3] := -0.26041505;
      FC_W[39,4] := 1.41878152;
      FC_W[39,5] := -1.64343119;
      FC_W[39,6] := -1.04960263;
      FC_W[39,7] := -2.64630604;
      FC_B[0] := 0.05778861;
      FC_B[1] := -0.77456111;
      FC_B[2] := 0.04080770;
      FC_B[3] := -0.51699263;
      FC_B[4] := -0.07885389;
      FC_B[5] := -0.07563572;
      FC_B[6] := 0.08624240;
      FC_B[7] := -0.51110834;
      FC_B[8] := -0.47873577;
      FC_B[9] := -0.51429105;
      FC_B[10] := -0.60357922;
      FC_B[11] := -0.94705731;
      FC_B[12] := -0.97999293;
      FC_B[13] := -1.39726925;
      FC_B[14] := 0.65040559;
      FC_B[15] := -0.85064948;
      FC_B[16] := 0.54259211;
      FC_B[17] := -0.08317784;
      FC_B[18] := 0.85150599;
      FC_B[19] := -1.14756417;
      FC_B[20] := -0.48967159;
      FC_B[21] := 0.13038819;
      FC_B[22] := -1.92337763;
      FC_B[23] := -1.60704899;
      FC_B[24] := -1.90559065;
      FC_B[25] := -1.90423548;
      FC_B[26] := -1.68349874;
      FC_B[27] := 0.44105780;
      FC_B[28] := 0.01162814;
      FC_B[29] := 1.81041276;
      FC_B[30] := -1.92445028;
      FC_B[31] := -1.91580296;
      FC_B[32] := -1.91381097;
      FC_B[33] := -1.90096831;
      FC_B[34] := -1.90703869;
      FC_B[35] := -1.90360427;
      FC_B[36] := -0.76133698;
      FC_B[37] := -1.89931357;
      FC_B[38] := 0.72174245;
      FC_B[39] := 0.76041430;

END_DATA_BLOCK
